            Script: movej(get_inverse_kin(pose_trans(FRM_Reference, PSE_A), qnear=JNT_Q), r=0.020)
          Else 
            Script: movej(pose_trans(FRM_Reference, PSE_A), r=0.020)
        MoveL speed 400 mm/s, acceleration 500 mm/s^2 (useActiveTCP=true) feature=FRM_Reference
          If PSE_T_H≠PSE_Z
            Waypoint Variable (Variable): motionParameters(blendRadius=0.01); variable=PSE_T_H
          Waypoint Variable (Variable): motionParameters(jointSpeed=1.047198 jointAcceleration=1.396263 cartesianSpeed=0.09 cartesianAcceleration=0.05); variable=PSE_T
            Until TOOL_CONTACT_DETECTION (allowActions=false retraction=NONE decelerationAcceleration=0.5 decelerationAngularAcceleration=34.906585)
          Force Frame feature=FRM_Reference; selection=[1, 1, 1, 0, 0, 0]; wrench=[0, 0, 0, 0, 0, 0]; limitsForce=[0.1, 0.1, 0.01, 1.047198, 1.047198, 1.047198]; limitsMotion=[0.1, 0.1, 0.1, 0.349066, 0.349066, 0.349066]
            Waypoint Variable (Variable): motionParameters(jointSpeed=1.047198 jointAcceleration=1.396263 cartesianSpeed=0.07 cartesianAcceleration=0.04); variable=PSE_T
          Folder EXTT
            Switch expression=JIG
              Case (caseValue=1)
                Folder 3FG
                  If OBJ_Picked
                    Set DigitalOutput pin=GRP_3F_Open; digitalValue=0
                    Wait Sleep waitTime=0.2
          Folder EOAT
            ''
    Case (caseValue=12)
      Folder Decap
        Action_Info := "decapping"
        Set DigitalOutput pin=GRP_3F_Enable; digitalValue=1
        Set DigitalOutput pin=GRP_3F_Decap; digitalValue=1
        Force Simple feature=Joint_6_name; selection=[0, 0, 1, 0, 0, 0]; wrench=[0, 0, 5, 0, 0, 0]; limitsForce=[0.15, 0.15, 0.15, 1.047198, 1.047198, 1.047198]; limitsMotion=[0.1, 0.1, 0.1, 0.349066, 0.349066, 0.349066]
          Script: check_decapping(offset=0.015, timeout=5, abort=CMD_Hold)
        Set DigitalOutput pin=GRP_3F_Decap; digitalValue=0
        Set DigitalOutput pin=GRP_3F_Enable; digitalValue=0
        MoveL speed 150 mm/s, acceleration 800 mm/s^2 (useActiveTCP=true) feature=FRM_Reference
          Waypoint Variable (Variable): variable=PSE_R
    Case (caseValue=13)
      Timer (action=Reset) variable(name=TMR_Barcode)
      Folder Read [hidden by the author, left out]
    Case (caseValue=15)
      Folder Detect
        Action_Info := "detect"
    Case (caseValue=30)
      Folder Shake
        Action_Info := "shake"
        Script: do_transition(pose_trans(FRM_Reference, PSE_T), keep_rxry=OBJ_Picked)
        If PSE_A_H≠PSE_Z
          If JNT_Q≠JNT_Z
            Script: movej(get_inverse_kin(pose_trans(FRM_Reference, PSE_A_H), qnear=JNT_Q), r=0.050)
          Else 
            Script: movej(pose_trans(FRM_Reference, PSE_A_H), r=0.050)
        If PSE_A≠PSE_Z
          If JNT_Q≠JNT_Z
            Script: movej(get_inverse_kin(pose_trans(FRM_Reference, PSE_A), qnear=JNT_Q), r=0.020)
          Else 
            Script: movej(pose_trans(FRM_Reference, PSE_A), r=0.020)
        MoveL speed 400 mm/s, acceleration 500 mm/s^2 (useActiveTCP=true) feature=FRM_Reference
          If PSE_T_H≠PSE_Z
            Waypoint Variable (Variable): motionParameters(blendRadius=0.01); variable=PSE_T_H
          Waypoint Variable (Variable): motionParameters(jointSpeed=1.047198 jointAcceleration=1.396263 cartesianSpeed=0.12 cartesianAcceleration=0.08); variable=PSE_T
          Folder EXTT
            ''
            MoveJ speed 60 deg/s, acceleration 80 deg/s^2 (useActiveTCP=true) feature=Base
              Waypoint Waypoint_6: TCP in base x=8.801 y=-547.927 z=402.697 mm, rx=-0.5899 ry=-0.0072 rz=-0.0613 rad; joints [-69.01, -76.872, -104.694, -56.634, 78.043, -158.781] deg; TCP offset x=0 y=0 z=161 mm, rx=3.1415 ry=0 rz=0 rad
            MoveJ speed 60 deg/s, acceleration 80 deg/s^2 (useActiveTCP=true) feature=Base
              Waypoint Waypoint_18: TCP in base x=-178.372 y=-433.927 z=368.082 mm, rx=-0.0866 ry=0.7047 rz=-0.0079 rad; joints [-72.502, -76.524, -102.817, -99.71, 50.308, -158.785] deg
            MoveJ speed 60 deg/s, acceleration 80 deg/s^2 (useActiveTCP=true) feature=Base
              Waypoint Waypoint_12: TCP in base x=8.801 y=-547.927 z=402.697 mm, rx=-0.5899 ry=-0.0072 rz=-0.0613 rad; joints [-69.01, -76.872, -104.694, -56.634, 78.043, -158.781] deg
            MoveJ speed 60 deg/s, acceleration 80 deg/s^2 (useActiveTCP=true) feature=Base
              Waypoint Waypoint_19: TCP in base x=-178.372 y=-433.927 z=368.082 mm, rx=-0.0866 ry=0.7047 rz=-0.0079 rad; joints [-72.502, -76.524, -102.817, -99.71, 50.308, -158.785] deg
          If PSE_R_H≠PSE_Z
            Waypoint Variable (Variable): motionParameters(blendRadius=0.01); variable=PSE_R
            Waypoint Variable (Variable): variable=PSE_R_H
          Else 
            Waypoint Variable (Variable): variable=PSE_R
    Case (caseValue=31)
      Action_Info := "Pick_Vial"
      Folder Pick_Vial
        URCap Gripper (Robotiq_Grippers, Robotiq Inc.) dataModel(position=0.0, force=27.84313725490196, speed=32.15686274509804, positionInDouble=0.0, forceInDouble=27.84313725490196, speedInDouble=32.15686274509804, slaveIds=[9], blocking=true)
        MoveJ speed 60 deg/s, acceleration 80 deg/s^2 (useActiveTCP=true) feature=Base
          Waypoint Vial_above: motionParameters(jointSpeed=0.436332 jointAcceleration=0.523599 cartesianSpeed=0.25 cartesianAcceleration=1.2 blendRadius=0.05); TCP in base x=17.106 y=-652.093 z=184.921 mm, rx=0 ry=0 rz=1.5641 rad; joints [-76.636, -112.403, -84.029, -73.556, 90.141, -256.27] deg
        MoveL speed 250 mm/s, acceleration 1200 mm/s^2 (useActiveTCP=true) feature=Base
          Waypoint Vial_pick_point: motionParameters(jointSpeed=1.047198 jointAcceleration=1.396263 cartesianSpeed=0.1 cartesianAcceleration=0.5); TCP in base x=17.106 y=-648.923 z=93.308 mm, rx=0 ry=0 rz=1.5641 rad; joints [-76.583, -116.742, -92.083, -61.164, 90.132, -256.177] deg
        URCap Gripper (Robotiq_Grippers, Robotiq Inc.) dataModel(position=100.0, force=32.94117647058823, speed=27.84313725490196, positionInDouble=100.0, forceInDouble=32.94117647058823, speedInDouble=27.84313725490196, slaveIds=[9], blocking=true)
        MoveL speed 250 mm/s, acceleration 1200 mm/s^2 (useActiveTCP=true) feature=Base
          Waypoint Waypoint_20: motionParameters(jointSpeed=1.047198 jointAcceleration=1.396263 cartesianSpeed=0.1 cartesianAcceleration=0.5 blendRadius=0.05); TCP in base x=19.228 y=-648.67 z=184.921 mm, rx=0 ry=0 rz=0.0241 rad; joints [-76.382, -111.96, -84.66, -73.372, 90.146, -167.779] deg
        SafeHome (positionOptionType=SPEED_AND_ACCELERATION speed=1.047198 acceleration=1.396263 nextMotionTime=2)
    Case (caseValue=32)
      decap := False
      Folder decap_Vial
        Set DigitalOutput pin=digital_out[5]; digitalValue=1
        MoveJ speed 60 deg/s, acceleration 80 deg/s^2 (useActiveTCP=true) feature=Base
          Waypoint Waypoint_33: motionParameters(jointSpeed=0.436332 jointAcceleration=0.523599 cartesianSpeed=0.25 cartesianAcceleration=1.2 blendRadius=0); TCP in base x=-32.362 y=-348.336 z=391.476 mm, rx=0 ry=0 rz=-0.0047 rad; joints [-72.819, -68.266, -97.918, -103.808, 90.124, -162.602] deg
        MoveL speed 250 mm/s, acceleration 1200 mm/s^2 (useActiveTCP=true) feature=Base
          Waypoint Vial_3FG_place: motionParameters(jointSpeed=1.047198 jointAcceleration=1.396263 cartesianSpeed=0.1 cartesianAcceleration=0.5); TCP in base x=-31.859 y=-349.403 z=145.301 mm, rx=0 ry=0 rz=0 rad; joints [-72.903, -71.756, -132.514, -65.722, 90.129, -162.805] deg
        Set DigitalOutput pin=digital_out[5]; digitalValue=0
        Wait Sleep waitTime=0.5
        MoveL speed 250 mm/s, acceleration 1200 mm/s^2 (useActiveTCP=true) feature=Base
          Waypoint Waypoint_34: motionParameters(jointSpeed=1.047198 jointAcceleration=1.396263 cartesianSpeed=0.1 cartesianAcceleration=0.5 blendRadius=0.05); TCP in base x=-32.362 y=-348.336 z=391.476 mm, rx=0 ry=0 rz=-0.0047 rad; joints [-72.819, -68.266, -97.918, -103.808, 90.124, -162.602] deg
        MoveJ speed 60 deg/s, acceleration 80 deg/s^2 (useActiveTCP=true) feature=Base
          Waypoint cap_dump: motionParameters(jointSpeed=0.436332 jointAcceleration=0.523599 cartesianSpeed=0.25 cartesianAcceleration=1.2); TCP in base x=-139.169 y=-420.164 z=146.096 mm, rx=0 ry=0 rz=0 rad; joints [-90.79, -86.479, -121, -62.513, 90.12, -180.712] deg
        URCap Gripper (Robotiq_Grippers, Robotiq Inc.) dataModel(position=0.0, force=100.0, speed=100.0, positionInDouble=0.0, forceInDouble=100.0, speedInDouble=100.0, slaveIds=[9], blocking=true)
        MoveJ speed 60 deg/s, acceleration 80 deg/s^2 (useActiveTCP=true) feature=Base
          Waypoint Waypoint_35: motionParameters(jointSpeed=0.436332 jointAcceleration=0.523599 cartesianSpeed=0.25 cartesianAcceleration=1.2 blendRadius=0.05); TCP in base x=-32.362 y=-348.336 z=391.476 mm, rx=0 ry=0 rz=-0.0047 rad; joints [-72.819, -68.266, -97.918, -103.808, 90.124, -162.602] deg
        MoveL speed 250 mm/s, acceleration 1200 mm/s^2 (useActiveTCP=true) feature=Base
          Waypoint Vial_3FG_place: motionParameters(jointSpeed=1.047198 jointAcceleration=1.396263 cartesianSpeed=0.1 cartesianAcceleration=0.5); TCP in base x=-31.859 y=-349.403 z=145.301 mm, rx=0 ry=0 rz=0 rad; joints [-72.903, -71.756, -132.514, -65.722, 90.129, -162.805] deg
        URCap Gripper (Robotiq_Grippers, Robotiq Inc.) dataModel(position=100.0, force=100.0, speed=80.0, positionInDouble=100.0, forceInDouble=100.0, speedInDouble=80.0, slaveIds=[9], blocking=true)
        SuppressedNode
          decap := True
        SuppressedNode
          Script: dynamic_upward_motion(0.015, 7)
        SuppressedNode
          MoveL speed 250 mm/s, acceleration 1200 mm/s^2 (useActiveTCP=true) feature=Joint_6_name
            MoveDirectionNode (selectedDirection=ZPlus toolParams=8.0E-4, 0.001) feature=Base
              Until DISTANCE (allowActions=false deceleration=3 distanceNodeType=STOP) Distance=0.01; motionParameters(blendRadius=0)
        SuppressedNode
          decap := False
        Folder Decap
          Action_Info := "decapping"
          Set DigitalOutput pin=GRP_3F_Enable; digitalValue=1
          Set DigitalOutput pin=GRP_3F_Decap; digitalValue=1
          Force Frame feature=Base; selection=[0, 0, 1, 0, 0, 0]; wrench=[0, 0, 1, 0, 0, 0]; limitsForce=[0.15, 0.15, 0.001, 1.047198, 1.047198, 1.047198]; limitsMotion=[0.1, 0.1, 0.1, 0.349066, 0.349066, 0.349066]
            Script: check_decapping(offset=0.015, timeout=10, abort=CMD_Hold)
          Set DigitalOutput pin=GRP_3F_Decap; digitalValue=0
          Set DigitalOutput pin=GRP_3F_Enable; digitalValue=0
          MoveL speed 250 mm/s, acceleration 1200 mm/s^2 (useActiveTCP=true) feature=Base
            Waypoint Waypoint_36: motionParameters(jointSpeed=1.047198 jointAcceleration=1.396263 cartesianSpeed=0.1 cartesianAcceleration=0.5 blendRadius=0.05); TCP in base x=-32.362 y=-348.336 z=391.476 mm, rx=0 ry=0 rz=-0.0047 rad; joints [-72.819, -68.266, -97.918, -103.808, 90.124, -162.602] deg
        MoveJ speed 60 deg/s, acceleration 80 deg/s^2 (useActiveTCP=true) feature=Base
          Waypoint cap_dump: motionParameters(jointSpeed=0.436332 jointAcceleration=0.523599 cartesianSpeed=0.25 cartesianAcceleration=1.2); TCP in base x=-139.169 y=-420.164 z=146.096 mm, rx=0 ry=0 rz=0 rad; joints [-90.79, -86.479, -121, -62.513, 90.12, -180.712] deg
        URCap Gripper (Robotiq_Grippers, Robotiq Inc.) dataModel(position=0.0, force=100.0, speed=80.0, positionInDouble=0.0, forceInDouble=100.0, speedInDouble=80.0, slaveIds=[9], blocking=true)
        MoveJ speed 60 deg/s, acceleration 80 deg/s^2 (useActiveTCP=true) feature=Base
          Waypoint Waypoint_37: motionParameters(jointSpeed=0.436332 jointAcceleration=0.523599 cartesianSpeed=0.25 cartesianAcceleration=1.2 blendRadius=0.036); TCP in base x=-32.362 y=-348.336 z=391.476 mm, rx=0 ry=0 rz=-0.0047 rad; joints [-72.819, -68.266, -97.918, -103.808, 90.124, -162.602] deg
    Case (caseValue=33)
      Folder Shake and liquid transfer
        MoveL speed 250 mm/s, acceleration 1200 mm/s^2 (useActiveTCP=true) feature=Base
          Waypoint Vial_liq_above: motionParameters(jointSpeed=1.047198 jointAcceleration=1.396263 cartesianSpeed=0.1 cartesianAcceleration=0.5); TCP in base x=-25.304 y=-338.759 z=426.628 mm, rx=-1.3159 ry=0.8 rz=-0.9283 rad; joints [-21.713, -86.8, -129.663, 45.096, -43.028, -184.708] deg
          Waypoint Vial_liq_pick_1: motionParameters(jointSpeed=1.047198 jointAcceleration=1.396263 cartesianSpeed=0.1 cartesianAcceleration=0.5); TCP in base x=-2.66 y=-335.985 z=159.39 mm, rx=-1.1505 ry=0.6732 rz=-1.0106 rad; joints [-20.975, -83.1, -137.831, -114.287, 46.064, -14.375] deg
          Waypoint Vial_liq_pick_2: motionParameters(jointSpeed=1.047198 jointAcceleration=1.396263 cartesianSpeed=0.1 cartesianAcceleration=0.5); TCP in base x=-41.402 y=-356.792 z=125.395 mm, rx=-1.1435 ry=0.6511 rz=-0.8787 rad; joints [-25.36, -82.348, -146.215, -101.788, 37.598, -24.648] deg
          URCap Gripper (Robotiq_Grippers, Robotiq Inc.) dataModel(position=100.0, force=27.84313725490196, speed=32.15686274509804, positionInDouble=100.0, forceInDouble=27.84313725490196, speedInDouble=32.15686274509804, slaveIds=[9], blocking=true)
          Wait Sleep waitTime=1
          Set DigitalOutput pin=digital_out[5]; digitalValue=1
          Wait Sleep waitTime=0.5
          Waypoint Vial_liq_above: motionParameters(jointSpeed=1.047198 jointAcceleration=1.396263 cartesianSpeed=0.05 cartesianAcceleration=0.3 blendRadius=0.05); TCP in base x=-25.304 y=-338.759 z=426.628 mm, rx=-1.3159 ry=0.8 rz=-0.9283 rad; joints [-21.713, -86.8, -129.663, 45.096, -43.028, -184.708] deg
        MoveL speed 250 mm/s, acceleration 1200 mm/s^2 (useActiveTCP=true) feature=Base
          Waypoint Liquid_midway: motionParameters(jointSpeed=1.047198 jointAcceleration=1.396263 cartesianSpeed=0.1 cartesianAcceleration=0.5 blendRadius=0); TCP in base x=57.575 y=-583.082 z=306.415 mm, rx=-1.3517 ry=0.1209 rz=-0.0969 rad; joints [-51.29, -97.606, -136.419, 36.185, 44.156, -168.768] deg
          Loop Counting (count=3) loopVariable(name=Loop_1)
            Waypoint shake_1: motionParameters(jointSpeed=1.047198 jointAcceleration=1.396263 cartesianSpeed=0.5 cartesianAcceleration=2); TCP in base x=57.575 y=-583.085 z=306.423 mm, rx=-1.361 ry=-0.1556 rz=-0.4381 rad; joints [-51.29, -97.606, -136.418, 36.185, 44.156, -145.5] deg
            Waypoint shake_2: motionParameters(jointSpeed=1.047198 jointAcceleration=1.396263 cartesianSpeed=0.5 cartesianAcceleration=2); TCP in base x=57.582 y=-583.091 z=306.44 mm, rx=-1.3088 ry=0.3685 rz=0.2149 rad; joints [-51.29, -97.606, -136.416, 36.185, 44.155, -190] deg
          Waypoint drop_above_1: motionParameters(jointSpeed=1.047198 jointAcceleration=1.396263 cartesianSpeed=0.1 cartesianAcceleration=0.5); TCP in base x=268.235 y=-467.784 z=226.22 mm, rx=-1.0278 ry=-0.4308 rz=1.0046 rad; joints [-53.609, -95.474, -138.959, 24.045, 105.829, -198.245] deg
          Waypoint drop_above_2: motionParameters(jointSpeed=1.047198 jointAcceleration=1.396263 cartesianSpeed=0.1 cartesianAcceleration=0.5); TCP in base x=219.042 y=-470.776 z=133.754 mm, rx=-0.313 ry=-0.3444 rz=1.5006 rad; joints [-60.743, -97.429, -119.175, -41.501, 111.324, -235.78] deg
          Waypoint liq_tran_1: motionParameters(jointSpeed=1.047198 jointAcceleration=1.396263 cartesianSpeed=0.05 cartesianAcceleration=0.5 blendRadius=0.008); TCP in base x=213.068 y=-469.567 z=100.231 mm, rx=0.2519 ry=0.2179 rz=1.5928 rad; joints [-44.631, -104.414, -106.819, -71.743, 78.886, -225.335] deg
          Wait Sleep waitTime=1
          Waypoint drop_above_2: motionParameters(jointSpeed=1.047198 jointAcceleration=1.396263 cartesianSpeed=0.1 cartesianAcceleration=0.5); TCP in base x=219.042 y=-470.776 z=133.754 mm, rx=-0.313 ry=-0.3444 rz=1.5006 rad; joints [-60.743, -97.429, -119.175, -41.501, 111.324, -235.78] deg
          Waypoint Waypoint_21: motionParameters(jointSpeed=1.047198 jointAcceleration=1.396263 cartesianSpeed=0.1 cartesianAcceleration=0.5); TCP in base x=187.119 y=-493.959 z=133.754 mm, rx=-0.313 ry=-0.3444 rz=1.5006 rad; joints [-65.422, -99.182, -116.519, -44.234, 112.218, -240.733] deg
          Waypoint liq_tran_2: motionParameters(jointSpeed=1.047198 jointAcceleration=1.396263 cartesianSpeed=0.05 cartesianAcceleration=0.5); TCP in base x=195.958 y=-493.023 z=100.231 mm, rx=0.1607 ry=0.1098 rz=1.5253 rad; joints [-50.52, -104.533, -106.862, -66.514, 83.832, -227.689] deg
          Wait Sleep waitTime=1
          Waypoint drop_above_2: motionParameters(jointSpeed=1.047198 jointAcceleration=1.396263 cartesianSpeed=0.1 cartesianAcceleration=0.5); TCP in base x=219.042 y=-470.776 z=133.754 mm, rx=-0.313 ry=-0.3444 rz=1.5006 rad; joints [-60.743, -97.429, -119.175, -41.501, 111.324, -235.78] deg
          Waypoint drop_above_1: motionParameters(jointSpeed=1.047198 jointAcceleration=1.396263 cartesianSpeed=0.1 cartesianAcceleration=0.5); TCP in base x=268.235 y=-467.784 z=226.22 mm, rx=-1.0278 ry=-0.4308 rz=1.0046 rad; joints [-53.609, -95.474, -138.959, 24.045, 105.829, -198.245] deg
          Waypoint Liquid_midway: motionParameters(jointSpeed=1.047198 jointAcceleration=1.396263 cartesianSpeed=0.1 cartesianAcceleration=0.5); TCP in base x=57.575 y=-583.082 z=306.415 mm, rx=-1.3517 ry=0.1209 rz=-0.0969 rad; joints [-51.29, -97.606, -136.419, 36.185, 44.156, -168.768] deg
        MoveL speed 250 mm/s, acceleration 1200 mm/s^2 (useActiveTCP=true) feature=Base
          Waypoint Vial_drop_above: motionParameters(jointSpeed=1.047198 jointAcceleration=1.396263 cartesianSpeed=0.1 cartesianAcceleration=0.5); TCP in base x=0.325 y=-648.57 z=221.894 mm, rx=-0.8735 ry=1.1659 rz=-1.4827 rad; joints [-60.601, -137.11, -52.92, -147.418, 45.283, -19.072] deg
          Waypoint Vial_liq_drop: motionParameters(jointSpeed=1.047198 jointAcceleration=1.396263 cartesianSpeed=0.1 cartesianAcceleration=0.5); TCP in base x=1.021 y=-647.66 z=92.916 mm, rx=-0.8348 ry=1.0819 rz=-1.5406 rad; joints [-60.917, -140.075, -64.676, -125.954, 46.582, -22.337] deg
          URCap Gripper (Robotiq_Grippers, Robotiq Inc.) dataModel(position=0.0, force=27.84313725490196, speed=32.15686274509804, positionInDouble=0.0, forceInDouble=27.84313725490196, speedInDouble=32.15686274509804, slaveIds=[9], blocking=true)
          Waypoint Vial_drop_above: motionParameters(jointSpeed=1.047198 jointAcceleration=1.396263 cartesianSpeed=0.1 cartesianAcceleration=0.5); TCP in base x=0.325 y=-648.57 z=221.894 mm, rx=-0.8735 ry=1.1659 rz=-1.4827 rad; joints [-60.601, -137.11, -52.92, -147.418, 45.283, -19.072] deg
    Case (caseValue=34)
      SafeHome (positionOptionType=SPEED_AND_ACCELERATION speed=1.047198 acceleration=1.396263 nextMotionTime=2)
      MoveJ speed 60 deg/s, acceleration 80 deg/s^2 (useActiveTCP=true) feature=Base
        Waypoint Waypoint_9: motionParameters(jointSpeed=0.436332 jointAcceleration=0.523599 cartesianSpeed=0.25 cartesianAcceleration=1.2); TCP in base x=206.301 y=-401.796 z=209.941 mm, rx=0 ry=0 rz=1.5608 rad; joints [-45.627, -84.145, -113.025, -72.821, 90.127, -225.014] deg
      MoveL speed 250 mm/s, acceleration 1200 mm/s^2 (useActiveTCP=true) feature=Base
        Waypoint Waypoint_10: motionParameters(jointSpeed=1.047198 jointAcceleration=1.396263 cartesianSpeed=0.1 cartesianAcceleration=0.5); TCP in base x=200.866 y=-400.818 z=105.073 mm, rx=0 ry=0 rz=1.5608 rad; joints [-46.083, -90.669, -123.933, -55.389, 90.105, -225.416] deg
      URCap Gripper (Robotiq_Grippers, Robotiq Inc.) dataModel(position=100.0, force=27.84313725490196, speed=32.15686274509804, positionInDouble=100.0, forceInDouble=27.84313725490196, speedInDouble=32.15686274509804, slaveIds=[9], blocking=true)
      Wait Sleep waitTime=1
      MoveL speed 250 mm/s, acceleration 1200 mm/s^2 (useActiveTCP=true) feature=Base
        Waypoint Waypoint_11: motionParameters(jointSpeed=1.047198 jointAcceleration=1.396263 cartesianSpeed=0.1 cartesianAcceleration=0.5 blendRadius=0.05); TCP in base x=200.866 y=-400.818 z=325.177 mm, rx=0 ry=0 rz=1.5608 rad; joints [-46.018, -81.306, -98.396, -90.289, 90.129, -225.47] deg
      MoveJ speed 60 deg/s, acceleration 80 deg/s^2 (useActiveTCP=true) feature=Base
        Waypoint Waypoint_7: motionParameters(jointSpeed=0.436332 jointAcceleration=0.523599 cartesianSpeed=0.25 cartesianAcceleration=1.2 blendRadius=0.05); TCP in base x=-615.829 y=233.809 z=300 mm, rx=0.0051 ry=0.0087 rz=-2.1118 rad; joints [-188.832, -110.936, -69.076, -89.912, 89.674, -157.919] deg
      MoveL speed 250 mm/s, acceleration 1200 mm/s^2 (useActiveTCP=true) feature=Base
        Waypoint Waypoint_8: motionParameters(jointSpeed=1.047198 jointAcceleration=1.396263 cartesianSpeed=0.1 cartesianAcceleration=0.5); TCP in base x=-615.829 y=233.809 z=13.91 mm, rx=0.0051 ry=0.0087 rz=-2.1118 rad; joints [-188.874, -123.68, -94.539, -51.707, 89.657, -157.833] deg
      URCap Gripper (Robotiq_Grippers, Robotiq Inc.) dataModel(position=0.0, force=27.84313725490196, speed=32.15686274509804, positionInDouble=0.0, forceInDouble=27.84313725490196, speedInDouble=32.15686274509804, slaveIds=[9], blocking=true)
      MoveJ speed 60 deg/s, acceleration 80 deg/s^2 (useActiveTCP=true) feature=Base
        Waypoint Waypoint_7: motionParameters(jointSpeed=0.436332 jointAcceleration=0.523599 cartesianSpeed=0.25 cartesianAcceleration=1.2); TCP in base x=-615.829 y=233.809 z=300 mm, rx=0.0051 ry=0.0087 rz=-2.1118 rad; joints [-188.832, -110.936, -69.076, -89.912, 89.674, -157.919] deg
      SafeHome (positionOptionType=SPEED_AND_ACCELERATION speed=1.047198 acceleration=1.396263 nextMotionTime=2)
      SuppressedNode
        Folder Decap
          Action_Info := "decapping"
          Set DigitalOutput pin=GRP_3F_Enable; digitalValue=1
          Set DigitalOutput pin=GRP_3F_Decap; digitalValue=1
          Force Frame feature=Base; selection=[0, 0, 1, 0, 0, 0]; wrench=[0, 0, 1, 0, 0, 0]; limitsForce=[0.15, 0.15, 0.001, 1.047198, 1.047198, 1.047198]; limitsMotion=[0.1, 0.1, 0.1, 0.349066, 0.349066, 0.349066]
            Script: check_decapping(offset=0.015, timeout=10, abort=CMD_Hold)
          Set DigitalOutput pin=GRP_3F_Decap; digitalValue=0
          Set DigitalOutput pin=GRP_3F_Enable; digitalValue=0
          MoveL speed 250 mm/s, acceleration 1200 mm/s^2 (useActiveTCP=true) feature=Base
            Waypoint Waypoint_5: motionParameters(jointSpeed=1.047198 jointAcceleration=1.396263 cartesianSpeed=0.1 cartesianAcceleration=0.5 blendRadius=0.05); TCP in base x=-31.859 y=-349.402 z=312.809 mm, rx=0 ry=0 rz=0 rad; joints [-72.832, -66.838, -110.376, -92.778, 90.139, -162.834] deg
          MoveJ speed 60 deg/s, acceleration 80 deg/s^2 (useActiveTCP=true) feature=Base
            Waypoint cap_dump: motionParameters(jointSpeed=0.436332 jointAcceleration=0.523599 cartesianSpeed=0.25 cartesianAcceleration=1.2); TCP in base x=-139.169 y=-420.164 z=146.096 mm, rx=0 ry=0 rz=0 rad; joints [-90.79, -86.479, -121, -62.513, 90.12, -180.712] deg
          URCap Gripper (Robotiq_Grippers, Robotiq Inc.) dataModel(position=0.0, force=100.0, speed=100.0, positionInDouble=0.0, forceInDouble=100.0, speedInDouble=100.0, slaveIds=[9], blocking=true)
          MoveJ speed 60 deg/s, acceleration 80 deg/s^2 (useActiveTCP=true) feature=Base
            Waypoint Waypoint_5: motionParameters(jointSpeed=0.436332 jointAcceleration=0.523599 cartesianSpeed=0.25 cartesianAcceleration=1.2 blendRadius=0.05); TCP in base x=-31.859 y=-349.402 z=312.809 mm, rx=0 ry=0 rz=0 rad; joints [-72.832, -66.838, -110.376, -92.778, 90.139, -162.834] deg
          Set DigitalOutput pin=digital_out[5]; digitalValue=1
    Case (caseValue=35)
      Folder Pick the powder container
        Wait Sleep waitTime=1
        MoveJ speed 60 deg/s, acceleration 80 deg/s^2 (useActiveTCP=true) feature=Base
          Waypoint Container_midwa: motionParameters(blendRadius=0.05); TCP in base x=-379.239 y=-127.191 z=300 mm, rx=0 ry=0 rz=-1.2472 rad; joints [-141.945, -74.312, -107.466, -88.214, 90.137, -160.485] deg
          Waypoint Container_capt: TCP in base x=-525.59 y=407.248 z=411.588 mm, rx=0 ry=0 rz=-2.8961 rad; joints [-206.083, -114.879, -46.847, -108.265, 90.132, -130.312] deg
        URCap VISOR Robotic App (SensoPart VISOR Robotic, SensoPart Industriesensorik GmbH) dataModel(visorAppTemplate=1); state(isChildrenLocked=true)
          URCap Easy Pick Setup (SensoPart VISOR Robotic, SensoPart Industriesensorik GmbH) dataModel(visorId=0, visorSetJob=true, visorJobName=Container_S, visorImageAcqSetup=2, visorCalibSetNo=7, visorDetector=1, visorImageAcqSource=1, visorOffsetSet=true, visorSetupStatus=3, Pose(key=visorImageAcqPose, Position(key=posePosition, Length(key=X value=-0.51041 unit=M), Length(key=Y value=0.417301 unit=M), Length(key=Z value=0.464095 unit=M)), Rotation(key=poseRotation, Angle(key=RX value=0.000026 unit=RAD), Angle(key=RY value=-0.000024 unit=RAD), Angle(key=RZ value=-2.896187 unit=RAD))), Pose(key=visorGripPose, Position(key=posePosition, Length(key=X value=-0.52891 unit=M), Length(key=Y value=0.461593 unit=M), Length(key=Z value=-0.178186 unit=M)), Rotation(key=poseRotation, Angle(key=RX value=-0.279814 unit=RAD), Angle(key=RY value=2.118244 unit=RAD), Angle(key=RZ value=-2.110314 unit=RAD)))); state(isChildrenLocked=true)
          URCap Process (SensoPart VISOR Robotic, SensoPart Industriesensorik GmbH) dataModel(Variable(key=visorCounterVar, variable(name=easyPickCount, initializeExpression=0)), Variable(key=visorPartsFoundVar, variable(name=easyPickParts, initializeExpression=0))); state(isChildrenLocked=true)
            URCap Image Acquisition Pose (SensoPart VISOR Robotic, SensoPart Industriesensorik GmbH) state(isChildrenLocked=true)
            URCap Object Detected (SensoPart VISOR Robotic, SensoPart Industriesensorik GmbH) state(isChildrenLocked=true)
              Folder Open Gripper
                URCap Gripper (Robotiq_Grippers, Robotiq Inc.) dataModel(position=0.0, force=30.0, speed=40.0, positionInDouble=0.0, forceInDouble=30.0, speedInDouble=40.0, slaveIds=[9], blocking=true)
                MoveJ speed 60 deg/s, acceleration 80 deg/s^2 (useActiveTCP=true) feature=Base
                  Waypoint Waypoint_13: TCP in base x=-479.451 y=284.141 z=125.27 mm, rx=-0.2768 ry=2.0984 rz=-2.1213 rad; joints [-165.671, -112.009, -127.874, -95.426, 1.192, -23.029] deg
              URCap Approach Pose (SensoPart VISOR Robotic, SensoPart Industriesensorik GmbH) dataModel(visorOffsetZ=-50.0); state(isChildrenLocked=true)
              URCap Target Pose (SensoPart VISOR Robotic, SensoPart Industriesensorik GmbH) state(isChildrenLocked=true)
              Folder Close Gripper
                URCap Gripper (Robotiq_Grippers, Robotiq Inc.) dataModel(position=100.0, force=30.19607843137255, speed=40.0, positionInDouble=100.0, forceInDouble=30.19607843137255, speedInDouble=40.0, slaveIds=[9], blocking=true)
              URCap Exit Pose (SensoPart VISOR Robotic, SensoPart Industriesensorik GmbH) dataModel(visorOffsetZ=-50.0); state(isChildrenLocked=true)
            URCap No Object Detected (SensoPart VISOR Robotic, SensoPart Industriesensorik GmbH) dataModel(Variable(key=visorNoObjCountVar, variable(name=easyPickNoObj, initializeExpression=0)))
              Popup Message (haltProgram=false message=No Container detected inputType=Text)
        MoveJ speed 60 deg/s, acceleration 80 deg/s^2 (useActiveTCP=true) feature=Base
          SuppressedNode
            Waypoint Cont_midwa_1: motionParameters(jointSpeed=1.047198 jointAcceleration=1.396263 cartesianSpeed=0.25 cartesianAcceleration=1.2 blendRadius=0.01); TCP in base x=-462.252 y=294.856 z=204.322 mm, rx=-0.3472 ry=2.0343 rz=-2.0655 rad; joints [-166.773, -128.859, -129.893, 70.604, 5.32, -171.145] deg
          Waypoint Waypoint_1: motionParameters(jointSpeed=0.523599 jointAcceleration=0.698132 cartesianSpeed=0.25 cartesianAcceleration=1.2 blendRadius=0); TCP in base x=-472.821 y=292.44 z=207.418 mm, rx=-0.2598 ry=-2.0535 rz=2.0707 rad; joints [-170.164, -118.699, -96.461, -142.976, 25.725, -0.32] deg
          Waypoint Waypoint_2: motionParameters(jointSpeed=0.523599 jointAcceleration=0.872665 cartesianSpeed=0.25 cartesianAcceleration=1.2 blendRadius=0.05); TCP in base x=-312.961 y=-152.991 z=223.61 mm, rx=-0.7453 ry=-1.7139 rz=1.6733 rad; joints [-134.992, -125.122, -83.555, -151.463, 94.666, 2.49] deg
          Waypoint Waypoint_3: motionParameters(jointSpeed=0.523599 jointAcceleration=0.698132 cartesianSpeed=0.25 cartesianAcceleration=1.2 blendRadius=0.05); TCP in base x=-113.75 y=-390.11 z=317.307 mm, rx=-0.5194 ry=-0.8399 rz=1.7569 rad; joints [-108.345, -98.585, -86.606, -121.699, 124.957, 41.411] deg
        MoveL speed 250 mm/s, acceleration 1200 mm/s^2 (useActiveTCP=true) feature=Base
          Waypoint Waypoint_15: motionParameters(jointSpeed=1.047198 jointAcceleration=1.396263 cartesianSpeed=0.1 cartesianAcceleration=0.5 blendRadius=0.05); TCP in base x=29.144 y=-436.802 z=327.885 mm, rx=-0.5216 ry=-0.6236 rz=1.8627 rad; joints [-89.657, -89.204, -96.411, -97.086, 128.129, 64.023] deg
          Waypoint Waypoint_14: motionParameters(jointSpeed=1.047198 jointAcceleration=1.396263 cartesianSpeed=0.1 cartesianAcceleration=0.3); TCP in base x=68.712 y=-569.42 z=285.215 mm, rx=-0.6792 ry=-0.7121 rz=1.394 rad; joints [-90.137, -103.3, -96.148, -70.007, 141.633, 93.932] deg
          Waypoint Waypoint_4: motionParameters(jointSpeed=1.047198 jointAcceleration=1.396263 cartesianSpeed=0.05 cartesianAcceleration=0.3); TCP in base x=-47.22 y=-557.625 z=136.371 mm, rx=-0.6792 ry=-0.7121 rz=1.394 rad; joints [-101.643, -114.727, -100.71, -68.127, 140.302, 75.797] deg
        URCap Gripper (Robotiq_Grippers, Robotiq Inc.) dataModel(position=0.0, force=30.0, speed=40.0, positionInDouble=0.0, forceInDouble=30.0, speedInDouble=40.0, slaveIds=[9], blocking=true)
        MoveL speed 250 mm/s, acceleration 1200 mm/s^2 (useActiveTCP=true) feature=Base
          Waypoint Waypoint_25: motionParameters(jointSpeed=1.047198 jointAcceleration=1.396263 cartesianSpeed=0.1 cartesianAcceleration=0.3); TCP in base x=65.436 y=-569.388 z=287.821 mm, rx=-0.6792 ry=-0.7121 rz=1.394 rad; joints [-90.466, -103.248, -95.699, -70.925, 141.635, 93.398] deg
          Waypoint Waypoint_15: motionParameters(jointSpeed=1.047198 jointAcceleration=1.396263 cartesianSpeed=0.1 cartesianAcceleration=0.5 blendRadius=0.05); TCP in base x=29.144 y=-436.802 z=327.885 mm, rx=-0.5216 ry=-0.6236 rz=1.8627 rad; joints [-89.657, -89.204, -96.411, -97.086, 128.129, 64.023] deg
        SafeHome (positionOptionType=SPEED_AND_ACCELERATION speed=1.047198 acceleration=1.396263 nextMotionTime=2)
        SuppressedNode
          MoveJ speed 60 deg/s, acceleration 80 deg/s^2 (useActiveTCP=true) feature=Base
            Waypoint Container_midwa: motionParameters(blendRadius=0.05); TCP in base x=-379.239 y=-127.191 z=300 mm, rx=0 ry=0 rz=-1.2472 rad; joints [-141.945, -74.312, -107.466, -88.214, 90.137, -160.485] deg
        URCap VISOR Robotic App (SensoPart VISOR Robotic, SensoPart Industriesensorik GmbH) dataModel(visorAppTemplate=1); state(isChildrenLocked=true)
          URCap Easy Pick Setup (SensoPart VISOR Robotic, SensoPart Industriesensorik GmbH) dataModel(visorId=0, visorSetJob=true, visorJobName=Target_container, visorImageAcqSetup=2, visorCalibSetNo=7, visorImageAcqSource=0, visorDetector=1, visorOffsetSet=true, visorSetupStatus=3, Pose(key=visorGripPose, Position(key=posePosition, Length(key=X value=-0.43018 unit=M), Length(key=Y value=0.500077 unit=M), Length(key=Z value=-0.155571 unit=M)), Rotation(key=poseRotation, Angle(key=RX value=0.000011 unit=RAD), Angle(key=RY value=0.000015 unit=RAD), Angle(key=RZ value=-2.896111 unit=RAD))), Pose(key=visorImageAcqPose, Position(key=posePosition, Length(key=X value=-0.391157 unit=M), Length(key=Y value=0.420635 unit=M), Length(key=Z value=0.411587 unit=M)), Rotation(key=poseRotation, Angle(key=RX value=-0.000006 unit=RAD), Angle(key=RY value=-0.000024 unit=RAD), Angle(key=RZ value=-2.896146 unit=RAD)))); state(isChildrenLocked=true)
          URCap Process (SensoPart VISOR Robotic, SensoPart Industriesensorik GmbH) dataModel(Variable(key=visorCounterVar, variable(name=easyPickCount_1, initializeExpression=0)), Variable(key=visorPartsFoundVar, variable(name=easyPickParts_1, initializeExpression=0))); state(isChildrenLocked=true)
            URCap Image Acquisition Pose (SensoPart VISOR Robotic, SensoPart Industriesensorik GmbH) state(isChildrenLocked=true)
            URCap Object Detected (SensoPart VISOR Robotic, SensoPart Industriesensorik GmbH) state(isChildrenLocked=true)
              Folder Open Gripper
                URCap Gripper (Robotiq_Grippers, Robotiq Inc.) dataModel(position=0.0, force=30.0, speed=40.0, positionInDouble=0.0, forceInDouble=30.0, speedInDouble=40.0, slaveIds=[9], blocking=true)
              URCap Approach Pose (SensoPart VISOR Robotic, SensoPart Industriesensorik GmbH) dataModel(visorOffsetZ=-50.0); state(isChildrenLocked=true)
              URCap Target Pose (SensoPart VISOR Robotic, SensoPart Industriesensorik GmbH) state(isChildrenLocked=true)
              Folder Close Gripper
                URCap Gripper (Robotiq_Grippers, Robotiq Inc.) dataModel(position=100.0, force=30.19607843137255, speed=40.0, positionInDouble=100.0, forceInDouble=30.19607843137255, speedInDouble=40.0, slaveIds=[9], blocking=true)
              URCap Exit Pose (SensoPart VISOR Robotic, SensoPart Industriesensorik GmbH) dataModel(visorOffsetZ=-50.0); state(isChildrenLocked=true)
            URCap No Object Detected (SensoPart VISOR Robotic, SensoPart Industriesensorik GmbH) dataModel(Variable(key=visorNoObjCountVar, variable(name=easyPickNoObj_1, initializeExpression=0)))
              Popup Message (haltProgram=false message=No Target container is detected inputType=Text)
        MoveJ speed 60 deg/s, acceleration 80 deg/s^2 (useActiveTCP=true) feature=Base
          Waypoint Waypoint_16: motionParameters(jointSpeed=0.698132 jointAcceleration=0.872665 cartesianSpeed=0.25 cartesianAcceleration=1.2); TCP in base x=-389.004 y=141.378 z=266.753 mm, rx=0.0001 ry=-0.0001 rz=-2.8961 rad; joints [-181.152, -76.776, -110.541, -82.676, 90.144, -105.201] deg
          Waypoint Waypoint_17: motionParameters(jointSpeed=0.698132 jointAcceleration=0.872665 cartesianSpeed=0.25 cartesianAcceleration=1.2); TCP in base x=-35.034 y=-360.271 z=346.67 mm, rx=0.0001 ry=0 rz=-1.4195 rad; joints [-73.886, -68.929, -104.178, -96.885, 90.142, -82.58] deg
        Set DigitalOutput pin=digital_out[5]; digitalValue=1
        MoveL speed 250 mm/s, acceleration 1200 mm/s^2 (useActiveTCP=true) feature=Base
          Waypoint Waypoint_22: motionParameters(jointSpeed=1.047198 jointAcceleration=1.396263 cartesianSpeed=0.1 cartesianAcceleration=0.5); TCP in base x=-31.771 y=-348.512 z=220.918 mm, rx=0.0001 ry=0 rz=-1.1964 rad; joints [-72.82, -67.691, -123.366, -78.936, 90.15, -94.217] deg
          Waypoint Waypoint_23: motionParameters(jointSpeed=1.047198 jointAcceleration=1.396263 cartesianSpeed=0.05 cartesianAcceleration=0.3); TCP in base x=-31.891 y=-348.193 z=178.714 mm, rx=0.0001 ry=0 rz=-1.1964 rad; joints [-72.841, -69.405, -128.724, -71.864, 90.145, -94.213] deg
        Set DigitalOutput pin=digital_out[5]; digitalValue=0
        Wait Sleep waitTime=1
        URCap Gripper (Robotiq_Grippers, Robotiq Inc.) dataModel(position=0.0, force=30.19607843137255, speed=40.0, positionInDouble=0.0, forceInDouble=30.19607843137255, speedInDouble=40.0, slaveIds=[9], blocking=true)
        MoveL speed 250 mm/s, acceleration 1200 mm/s^2 (useActiveTCP=true) feature=Base
          Waypoint Waypoint_24: motionParameters(jointSpeed=1.047198 jointAcceleration=1.396263 cartesianSpeed=0.05 cartesianAcceleration=0.3); TCP in base x=-31.773 y=-348.52 z=270.997 mm, rx=0.0001 ry=0 rz=-1.1964 rad; joints [-72.799, -66.725, -116.549, -86.72, 90.151, -94.226] deg
        SafeHome (positionOptionType=SPEED_AND_ACCELERATION speed=1.047198 acceleration=1.396263 nextMotionTime=2)
    Case (caseValue=36)
      MoveL speed 250 mm/s, acceleration 1200 mm/s^2 (useActiveTCP=true) feature=Base
        Waypoint Waypoint_26: TCP in base x=-30.182 y=-347.336 z=210.998 mm, rx=0 ry=0 rz=0 rad; joints [-72.486, -67.792, -124.787, -77.413, 90.141, -162.427] deg
      URCap Gripper (Robotiq_Grippers, Robotiq Inc.) dataModel(position=100.0, force=30.19607843137255, speed=40.0, positionInDouble=100.0, forceInDouble=30.19607843137255, speedInDouble=40.0, slaveIds=[9], blocking=true)
      Folder Decap
        Action_Info := "decapping"
        Set DigitalOutput pin=GRP_3F_Enable; digitalValue=1
        Set DigitalOutput pin=GRP_3F_Decap; digitalValue=1
        Force Frame feature=Base; selection=[0, 0, 1, 0, 0, 0]; wrench=[0, 0, 1, 0, 0, 0]; limitsForce=[0.15, 0.15, 0.001, 1.047198, 1.047198, 1.047198]; limitsMotion=[0.1, 0.1, 0.1, 0.349066, 0.349066, 0.349066]
          Script: check_decapping(offset=0.015, timeout=12, abort=CMD_Hold)
        Set DigitalOutput pin=GRP_3F_Decap; digitalValue=0
        Set DigitalOutput pin=GRP_3F_Enable; digitalValue=0
        MoveL speed 250 mm/s, acceleration 1200 mm/s^2 (useActiveTCP=true) feature=Base
          Waypoint Waypoint_27: motionParameters(jointSpeed=1.047198 jointAcceleration=1.396263 cartesianSpeed=0.1 cartesianAcceleration=0.5 blendRadius=0.05); TCP in base x=-30.361 y=-347.415 z=279.539 mm, rx=0 ry=0 rz=-0.0004 rad; joints [-72.488, -66.465, -115.449, -88.079, 90.139, -162.449] deg
          Waypoint Waypoint_28: motionParameters(jointSpeed=1.047198 jointAcceleration=1.396263 cartesianSpeed=0.1 cartesianAcceleration=0.5 blendRadius=0.05); TCP in base x=-154.725 y=-473.257 z=246.189 mm, rx=0 ry=0 rz=-0.0004 rad; joints [-92.526, -89.454, -102.579, -77.959, 90.132, -182.495] deg
          Waypoint Waypoint_29: motionParameters(jointSpeed=1.047198 jointAcceleration=1.396263 cartesianSpeed=0.1 cartesianAcceleration=0.3); TCP in base x=-145.695 y=-485.909 z=46.677 mm, rx=0 ry=0 rz=-0.0004 rad; joints [-91.444, -104.036, -119.144, -46.812, 90.094, -181.324] deg
        URCap Gripper (Robotiq_Grippers, Robotiq Inc.) dataModel(position=61.24306326304106, force=30.19607843137255, speed=40.0, positionInDouble=61.24306326304106, forceInDouble=30.19607843137255, speedInDouble=40.0, slaveIds=[9], blocking=true)
        MoveL speed 250 mm/s, acceleration 1200 mm/s^2 (useActiveTCP=true) feature=Base
          Waypoint Waypoint_38: motionParameters(jointSpeed=1.047198 jointAcceleration=1.396263 cartesianSpeed=0.1 cartesianAcceleration=0.5 blendRadius=0.05); TCP in base x=-145.695 y=-485.909 z=261.43 mm, rx=0 ry=0 rz=-0.0004 rad; joints [-91.4, -90.37, -99.399, -80.223, 90.132, -181.38] deg
          Waypoint Waypoint_30: motionParameters(jointSpeed=1.047198 jointAcceleration=1.396263 cartesianSpeed=0.1 cartesianAcceleration=0.5 blendRadius=0.05); TCP in base x=-30.182 y=-347.336 z=265.578 mm, rx=0 ry=0 rz=0 rad; joints [-72.462, -66.558, -117.437, -85.997, 90.142, -162.436] deg
          Waypoint Waypoint_31: motionParameters(jointSpeed=1.047198 jointAcceleration=1.396263 cartesianSpeed=0.1 cartesianAcceleration=0.5); TCP in base x=-30.182 y=-347.336 z=175.833 mm, rx=0 ry=0 rz=0 rad; joints [-72.5, -69.38, -129.182, -71.43, 90.136, -162.42] deg
        URCap Gripper (Robotiq_Grippers, Robotiq Inc.) dataModel(position=43.04106548279689, force=30.19607843137255, speed=40.0, positionInDouble=43.04106548279689, forceInDouble=30.19607843137255, speedInDouble=40.0, slaveIds=[9], blocking=true)
        Wait Sleep waitTime=1
        Set DigitalOutput pin=digital_out[5]; digitalValue=1
        MoveL speed 250 mm/s, acceleration 1200 mm/s^2 (useActiveTCP=true) feature=Base
          Waypoint Waypoint_32: motionParameters(jointSpeed=1.047198 jointAcceleration=1.396263 cartesianSpeed=0.1 cartesianAcceleration=0.5 blendRadius=0.05); TCP in base x=-30.182 y=-347.336 z=316.067 mm, rx=0 ry=0 rz=0 rad; joints [-72.438, -66.521, -110.081, -93.39, 90.138, -162.442] deg
        URCap VISOR Robotic App (SensoPart VISOR Robotic, SensoPart Industriesensorik GmbH) dataModel(visorAppTemplate=1); state(isChildrenLocked=true)
          URCap Easy Pick Setup (SensoPart VISOR Robotic, SensoPart Industriesensorik GmbH) dataModel(visorId=0, visorSetJob=true, visorJobName=Weigh_scale, visorImageAcqSetup=2, visorImageAcqSource=1, visorCalibSetNo=9, visorDetector=1, visorSetupStatus=5, visorOffsetSet=true, Pose(key=visorGripPose, Position(key=posePosition, Length(key=X value=-0.66092 unit=M), Length(key=Y value=-0.026261 unit=M), Length(key=Z value=0.113423 unit=M)), Rotation(key=poseRotation, Angle(key=RX value=0.044036 unit=RAD), Angle(key=RY value=-0.006733 unit=RAD), Angle(key=RZ value=-1.658906 unit=RAD)))); state(isChildrenLocked=true)
          URCap Process (SensoPart VISOR Robotic, SensoPart Industriesensorik GmbH) dataModel(Variable(key=visorCounterVar, variable(name=easyPickCount_2, initializeExpression=0)), Variable(key=visorPartsFoundVar, variable(name=easyPickParts_2, initializeExpression=0))); state(isChildrenLocked=true)
            URCap Image Acquisition Pose (SensoPart VISOR Robotic, SensoPart Industriesensorik GmbH) state(isChildrenLocked=true)
            URCap Object Detected (SensoPart VISOR Robotic, SensoPart Industriesensorik GmbH) state(isChildrenLocked=true)
              Folder Open Gripper
                Wait NoWait
              URCap Approach Pose (SensoPart VISOR Robotic, SensoPart Industriesensorik GmbH) dataModel(visorOffsetZ=-50.0); state(isChildrenLocked=true)
              URCap Target Pose (SensoPart VISOR Robotic, SensoPart Industriesensorik GmbH) state(isChildrenLocked=true)
              Folder Close Gripper
                URCap Gripper (Robotiq_Grippers, Robotiq Inc.) dataModel(position=0.0, force=30.19607843137255, speed=40.0, positionInDouble=0.0, forceInDouble=30.19607843137255, speedInDouble=40.0, slaveIds=[9], blocking=true)
              URCap Exit Pose (SensoPart VISOR Robotic, SensoPart Industriesensorik GmbH) dataModel(visorOffsetZ=-100.0); state(isChildrenLocked=true)
            URCap No Object Detected (SensoPart VISOR Robotic, SensoPart Industriesensorik GmbH) dataModel(Variable(key=visorNoObjCountVar, variable(name=easyPickNoObj_2, initializeExpression=0)))
              Popup Message (haltProgram=false message=No weigh scale is detected inputType=Text)
        SafeHome (positionOptionType=SPEED_AND_ACCELERATION speed=1.047198 acceleration=1.396263 nextMotionTime=2)
        MoveJ speed 60 deg/s, acceleration 80 deg/s^2 (useActiveTCP=true) feature=Base
          Waypoint Waypoint_39: TCP in base x=137.772 y=-577.76 z=300 mm, rx=0 ry=0 rz=-1.5944 rad; joints [-63.54, -101.785, -81.001, -87.198, 90.144, -62.245] deg
        MoveL speed 250 mm/s, acceleration 1200 mm/s^2 (useActiveTCP=true) feature=Base
          Waypoint Waypoint_41: motionParameters(jointSpeed=1.047198 jointAcceleration=1.396263 cartesianSpeed=0.1 cartesianAcceleration=0.5); TCP in base x=74.223 y=-565.642 z=234.62 mm, rx=-0.5169 ry=0.5292 rz=-1.5296 rad; joints [-54.985, -107.527, -85.329, -102.066, 60.279, -46.981] deg
          Waypoint Waypoint_40: motionParameters(jointSpeed=1.047198 jointAcceleration=1.396263 cartesianSpeed=0.05 cartesianAcceleration=0.3); TCP in base x=39.988 y=-564.833 z=191.055 mm, rx=-0.7676 ry=0.3431 rz=-2.2413 rad; joints [-57.701, -107.406, -92.471, -93.607, 59.17, -6.639] deg
        URCap Gripper (Robotiq_Grippers, Robotiq Inc.) dataModel(position=100.0, force=20.0, speed=30.0, positionInDouble=100.0, forceInDouble=20.0, speedInDouble=30.0, slaveIds=[9], blocking=true)
        Loop Counting (count=2) loopVariable(name=Loop_2)
          MoveL speed 250 mm/s, acceleration 1200 mm/s^2 (useActiveTCP=true) feature=Base
            Waypoint Waypoint_42: motionParameters(jointSpeed=1.047198 jointAcceleration=1.396263 cartesianSpeed=0.5 cartesianAcceleration=1.2 blendRadius=0); TCP in base x=41.363 y=-564.865 z=192.806 mm, rx=0.2785 ry=0.6241 rz=0.7623 rad; joints [-57.586, -107.397, -92.198, -93.963, 59.209, -186.442] deg
            Waypoint Waypoint_43: TCP in base x=41.363 y=-564.865 z=192.806 mm, rx=0.9734 ry=0.0641 rz=2.8083 rad; joints [-57.585, -107.391, -92.207, -93.949, 59.207, -310.817] deg
          URCap Gripper (Robotiq_Grippers, Robotiq Inc.) dataModel(position=24.83906770255271, force=20.0, speed=30.19607843137255, positionInDouble=24.83906770255271, forceInDouble=20.0, speedInDouble=30.19607843137255, slaveIds=[9], blocking=true)
          MoveL speed 250 mm/s, acceleration 1200 mm/s^2 (useActiveTCP=true) feature=Base
            Waypoint Waypoint_44: motionParameters(jointSpeed=1.047198 jointAcceleration=1.396263 cartesianSpeed=0.5 cartesianAcceleration=1.2 blendRadius=0); TCP in base x=40.883 y=-564.854 z=192.194 mm, rx=0.1109 ry=0.6592 rz=0.2757 rad; joints [-57.626, -107.402, -92.291, -93.842, 59.196, -157.494] deg
            Waypoint Waypoint_45: TCP in base x=42.648 y=-564.896 z=194.439 mm, rx=-0.4517 ry=0.5632 rz=-1.3434 rad; joints [-57.484, -107.381, -91.951, -94.273, 59.256, -60.779] deg
          URCap Gripper (Robotiq_Grippers, Robotiq Inc.) dataModel(position=78.43137254901961, force=20.0, speed=30.0, positionInDouble=78.43137254901961, forceInDouble=20.0, speedInDouble=30.0, slaveIds=[9], blocking=true)
        MoveL speed 250 mm/s, acceleration 1200 mm/s^2 (useActiveTCP=true) feature=Base
          Waypoint Waypoint_46: motionParameters(jointSpeed=1.047198 jointAcceleration=1.396263 cartesianSpeed=0.05 cartesianAcceleration=0.3); TCP in base x=99.944 y=-566.244 z=267.343 mm, rx=-0.4517 ry=0.5632 rz=-1.3434 rad; joints [-53.041, -108.287, -79.23, -108.385, 61.102, -56.184] deg
          Waypoint Waypoint_47: motionParameters(jointSpeed=1.047198 jointAcceleration=1.396263 cartesianSpeed=0.1 cartesianAcceleration=0.5 blendRadius=0); TCP in base x=99.944 y=-566.244 z=267.343 mm, rx=-0.1017 ry=0.0587 rz=-1.4579 rad; joints [-63.671, -99.121, -88.981, -82.751, 84.056, -70.038] deg
          Waypoint Waypoint_48: motionParameters(jointSpeed=1.047198 jointAcceleration=1.396263 cartesianSpeed=0.25 cartesianAcceleration=1.2); TCP in base x=-136.183 y=-647.487 z=294.248 mm, rx=-0.1017 ry=0.0587 rz=-1.4579 rad; joints [-87.788, -109.526, -72.49, -86.263, 84.243, -94.331] deg
          Waypoint Waypoint_49: TCP in base x=-159.024 y=-641.021 z=47.692 mm, rx=0 ry=0 rz=-1.4579 rad; joints [-92.238, -121.266, -92.571, -56.15, 90.14, -98.675] deg
        URCap Gripper (Robotiq_Grippers, Robotiq Inc.) dataModel(position=33.9400665926748, force=20.0, speed=30.19607843137255, positionInDouble=33.9400665926748, forceInDouble=20.0, speedInDouble=30.19607843137255, slaveIds=[9], blocking=true)
        MoveL speed 250 mm/s, acceleration 1200 mm/s^2 (useActiveTCP=true) feature=Base
          Waypoint Waypoint_50: TCP in base x=-159.024 y=-641.021 z=291.114 mm, rx=0 ry=0 rz=-1.4579 rad; joints [-92.2, -111.308, -69.838, -88.841, 90.151, -98.75] deg
          SafeHome (positionOptionType=SPEED_AND_ACCELERATION speed=1.047198 acceleration=1.396263 nextMotionTime=2)
    Case (caseValue=37)
      URCap VISOR Robotic App (SensoPart VISOR Robotic, SensoPart Industriesensorik GmbH) dataModel(visorAppTemplate=1); state(isChildrenLocked=true)
        URCap Easy Pick Setup (SensoPart VISOR Robotic, SensoPart Industriesensorik GmbH) dataModel(visorId=0, visorSetJob=true, visorJobName=Spatula, visorImageAcqSetup=2, visorImageAcqSource=1, visorCalibSetNo=10, visorDetector=1, visorSetupStatus=5, visorOffsetSet=true, Pose(key=visorGripPose, Position(key=posePosition, Length(key=X value=-0.650651 unit=M), Length(key=Y value=-0.390239 unit=M), Length(key=Z value=0.139774 unit=M)), Rotation(key=poseRotation, Angle(key=RX value=0.000035 unit=RAD), Angle(key=RY value=0.000024 unit=RAD), Angle(key=RZ value=2.990013 unit=RAD)))); state(isChildrenLocked=true)
        URCap Process (SensoPart VISOR Robotic, SensoPart Industriesensorik GmbH) dataModel(Variable(key=visorCounterVar, variable(name=easyPickCount_3, initializeExpression=0)), Variable(key=visorPartsFoundVar, variable(name=easyPickParts_3, initializeExpression=0))); state(isChildrenLocked=true)
          URCap Image Acquisition Pose (SensoPart VISOR Robotic, SensoPart Industriesensorik GmbH) state(isChildrenLocked=true)
          URCap Object Detected (SensoPart VISOR Robotic, SensoPart Industriesensorik GmbH) state(isChildrenLocked=true)
            Folder Open Gripper
              URCap Gripper (Robotiq_Grippers, Robotiq Inc.) dataModel(position=0.0, force=20.0, speed=30.19607843137255, positionInDouble=0.0, forceInDouble=20.0, speedInDouble=30.19607843137255, slaveIds=[9], blocking=true)
            URCap Approach Pose (SensoPart VISOR Robotic, SensoPart Industriesensorik GmbH) dataModel(visorOffsetZ=-100.0); state(isChildrenLocked=true)
            URCap Target Pose (SensoPart VISOR Robotic, SensoPart Industriesensorik GmbH) state(isChildrenLocked=true)
            Folder Close Gripper
              URCap Gripper (Robotiq_Grippers, Robotiq Inc.) dataModel(position=100.0, force=20.0, speed=30.19607843137255, positionInDouble=100.0, forceInDouble=20.0, speedInDouble=30.19607843137255, slaveIds=[9], blocking=true)
            URCap Exit Pose (SensoPart VISOR Robotic, SensoPart Industriesensorik GmbH) dataModel(visorOffsetZ=-250.0, visorToolSpeed=100.0, visorToolAcc=300.0); state(isChildrenLocked=true)
          URCap No Object Detected (SensoPart VISOR Robotic, SensoPart Industriesensorik GmbH) dataModel(Variable(key=visorNoObjCountVar, variable(name=easyPickNoObj_3, initializeExpression=0)))
            Popup Message (haltProgram=false message=No spatula is detected inputType=Text)
      MoveJ speed 60 deg/s, acceleration 80 deg/s^2 (useActiveTCP=true) feature=Base
        Waypoint Waypoint_51: motionParameters(jointSpeed=0.698132 jointAcceleration=0.872665 cartesianSpeed=0.25 cartesianAcceleration=1.2); TCP in base x=-138.513 y=-390.318 z=390.027 mm, rx=0.9851 ry=0.0766 rz=2.8273 rad; joints [-66.551, -74.061, -98.345, -115.037, 55.353, 37.764] deg
        Waypoint Waypoint_52: motionParameters(jointSpeed=0.698132 jointAcceleration=0.872665 cartesianSpeed=0.25 cartesianAcceleration=1.2); TCP in base x=200.663 y=-570.117 z=330.074 mm, rx=1.3605 ry=0.0217 rz=2.6816 rad; joints [-43.944, -124.326, -49.615, -141.861, 58.428, 68.113] deg
      MoveL speed 50 mm/s, acceleration 300 mm/s^2 (useActiveTCP=true) feature=Base
        Waypoint Waypoint_53: motionParameters(jointSpeed=1.047198 jointAcceleration=1.396263 cartesianSpeed=0.05 cartesianAcceleration=0.3); TCP in base x=200.65 y=-570.239 z=330.084 mm, rx=1.3605 ry=0.0217 rz=2.6816 rad; joints [-43.952, -124.342, -49.589, -141.868, 58.423, 68.107] deg
        Waypoint Waypoint_54: motionParameters(jointSpeed=1.047198 jointAcceleration=1.396263 cartesianSpeed=0.05 cartesianAcceleration=0.3); TCP in base x=143.03 y=-569.853 z=275.754 mm, rx=1.2979 ry=0.0264 rz=2.7129 rad; joints [-47.784, -117.454, -67.716, -126.008, 56.917, 63.329] deg
        Loop Counting (count=3) loopVariable(name=Loop_3)
          Waypoint Waypoint_55: motionParameters(jointSpeed=1.047198 jointAcceleration=1.396263 cartesianSpeed=0.05 cartesianAcceleration=0.3); TCP in base x=73.857 y=-577.013 z=221.505 mm, rx=1.2979 ry=0.0264 rz=2.7129 rad; joints [-52.913, -114.774, -80.289, -113.397, 53.656, 58.584] deg
            Until TOOL_CONTACT_DETECTION (allowActions=false retraction=0 decelerationAcceleration=3 decelerationAngularAcceleration=34.906585)
          Waypoint Waypoint_56: motionParameters(jointSpeed=1.047198 jointAcceleration=1.396263 cartesianSpeed=0.05 cartesianAcceleration=0.3); TCP in base x=135.677 y=-579.448 z=242.231 mm, rx=1.5554 ry=0.0154 rz=2.5559 rad; joints [-47.427, -124.812, -65.265, -134.284, 52.841, 72.036] deg
        Loop Counting (count=2) loopVariable(name=Loop_5)
          Waypoint Waypoint_56: motionParameters(jointSpeed=1.047198 jointAcceleration=1.396263 cartesianSpeed=0.05 cartesianAcceleration=0.3); TCP in base x=135.677 y=-579.448 z=242.231 mm, rx=1.5554 ry=0.0154 rz=2.5559 rad; joints [-47.427, -124.812, -65.265, -134.284, 52.841, 72.036] deg
          Waypoint Waypoint_57: motionParameters(jointSpeed=1.047198 jointAcceleration=1.396263 cartesianSpeed=0.5 cartesianAcceleration=1.2); TCP in base x=143.391 y=-581.809 z=226.065 mm, rx=1.6397 ry=0.0079 rz=2.5024 rad; joints [-46.773, -128.399, -63.349, -137.511, 52.317, 75.293] deg
        Waypoint Waypoint_59: motionParameters(jointSpeed=1.047198 jointAcceleration=1.396263 cartesianSpeed=0.05 cartesianAcceleration=0.3); TCP in base x=272.401 y=-578.183 z=239.561 mm, rx=2.127 ry=0.1139 rz=2.1556 rad; joints [-37.816, -154.733, -25.502, -178.522, 53.445, 96.624] deg
        Waypoint Waypoint_58: motionParameters(jointSpeed=1.047198 jointAcceleration=1.396263 cartesianSpeed=0.05 cartesianAcceleration=0.3); TCP in base x=223.649 y=-578.478 z=276.546 mm, rx=2.1743 ry=-0.0441 rz=2.0587 rad; joints [-41.771, -153.265, -25.455, -184.54, 55.381, 96.631] deg
      MoveJ speed 30 deg/s, acceleration 50 deg/s^2 (useActiveTCP=true) feature=Base
        Waypoint Waypoint_60: motionParameters(jointSpeed=0.349066 jointAcceleration=0.523599 cartesianSpeed=0.25 cartesianAcceleration=1.2 blendRadius=0.05); TCP in base x=-13.316 y=-544.772 z=383.372 mm, rx=2.2082 ry=0.0375 rz=2.0976 rad; joints [-53.447, -120.321, -68.514, -175.377, 39.556, 98.101] deg
        Waypoint Waypoint_61: motionParameters(jointSpeed=0.349066 jointAcceleration=0.523599 cartesianSpeed=0.25 cartesianAcceleration=1.2 blendRadius=0.05); TCP in base x=-412.189 y=-356.447 z=383.372 mm, rx=1.7517 ry=-0.74 rz=1.6007 rad; joints [-101.195, -120.321, -68.514, -175.377, 39.556, 98.101] deg
        Waypoint Waypoint_62: motionParameters(jointSpeed=0.349066 jointAcceleration=0.523599 cartesianSpeed=0.25 cartesianAcceleration=1.2); TCP in base x=-542.659 y=-114.282 z=251.262 mm, rx=1.813 ry=-0.6794 rz=1.6553 rad; joints [-123.661, -111.262, -103.952, -159.22, 12.548, 108.767] deg
      MoveL speed 250 mm/s, acceleration 1200 mm/s^2 (useActiveTCP=true) feature=Base
        Waypoint Waypoint_63: motionParameters(jointSpeed=1.047198 jointAcceleration=1.396263 cartesianSpeed=0.05 cartesianAcceleration=0.3); TCP in base x=-532.496 y=-127.81 z=159.342 mm, rx=1.813 ry=-0.6794 rz=1.6553 rad; joints [-121.654, -119.526, -108.357, -144.665, 14.532, 106.823] deg
        Waypoint Waypoint_64: motionParameters(jointSpeed=1.047198 jointAcceleration=1.396263 cartesianSpeed=0.05 cartesianAcceleration=0.3); TCP in base x=-576.035 y=-66.27 z=306.74 mm, rx=0.8621 ry=-0.2554 rz=2.1952 rad; joints [-142.141, -87.685, -107.535, -64.498, 50.077, -8.596] deg
        Waypoint Waypoint_65: motionParameters(jointSpeed=1.047198 jointAcceleration=1.396263 cartesianSpeed=0.05 cartesianAcceleration=0.3); TCP in base x=-581.965 y=-59.291 z=312.082 mm, rx=0.8621 ry=-0.2554 rz=2.1952 rad; joints [-143.275, -88.018, -106.65, -64.116, 50.29, -10.05] deg
        Waypoint Waypoint_66: motionParameters(jointSpeed=1.047198 jointAcceleration=1.396263 cartesianSpeed=0.5 cartesianAcceleration=1.2); TCP in base x=-581.965 y=-59.291 z=290.576 mm, rx=0.8621 ry=-0.2554 rz=2.1952 rad; joints [-143.281, -88.87, -109.094, -60.824, 50.286, -10.043] deg
        Waypoint Waypoint_67: TCP in base x=-581.965 y=-59.291 z=350.142 mm, rx=1.7575 ry=-0.6778 rz=1.6965 rad; joints [-131.863, -101.687, -97.87, -162.913, 4.302, 96.426] deg
      MoveJ speed 60 deg/s, acceleration 80 deg/s^2 (useActiveTCP=true) feature=Base
        Waypoint Waypoint_68: TCP in base x=-333.293 y=-480.744 z=350.142 mm, rx=2.2175 ry=0.1409 rz=2.2091 rad; joints [-82.414, -101.687, -97.87, -162.913, 4.302, 96.426] deg
  '=========='
  Folder PostSettings [hidden by the author, left out]
